// Geprüfte Kopie des aktiven Biegeplans. Schreibt nur FB_PlanStore, liest FB_BendKinematics und FB_BendSequence.
{attribute 'qualified_only'}
VAR_GLOBAL
    stActive : ST_PlanTransfer;
    bValid   : BOOL;
END_VAR

(* stored: Version 1.1.0.1
   GVL GVL_Plan: Id {e3de924e-5bdb-5771-a4f4-c570fdb85676} *)
